Fanuc KAREL source: kx00007.KL

-- PROVISIONAL review KL for V770-1; original PC SHA256 dfda3f059b3d32d90e934d8d872130bb282927e6442b5eb72e65107867753797
-- Incomplete behavior may be omitted. Consult companion uncertainty JSON. Do not deploy.
PROGRAM KX00007
%NOLOCKGROUP
VAR
  I : INTEGER
  J : INTEGER
  B : BOOLEAN
  F : FILE
  S : STRING[80]
-- UNRESOLVED_DECL P type=000102
BEGIN
  -- UNRESOLVED_PC offsets 5-13; opcodes 9D,2E,1F
  -- UNRESOLVED_PC offsets 18-22; opcodes 7F
END KX00007
